Fanuc KAREL source: kc00033.KL

-- PROVISIONAL review KL for V940-1; original PC SHA256 2e3bb30ba8f1449926ae04295cef8963f4468ff0dde0fae508bc08914172abd9
-- Incomplete behavior may be omitted. Consult companion uncertainty JSON. Do not deploy.
PROGRAM KC00033
%NOLOCKGROUP
BEGIN
  -- V9_ZERO_TABLE_METADATA_HINT layout=0001; no indexed target words; source/name/runtime held
  -- UNRESOLVED_PC offsets 5-32; opcodes 27,22,1C,22,22,76
  -- UNRESOLVED_PC offsets 37-41; opcodes 7F
END KC00033
